RoboDK station: Robot_3_2026.rdk

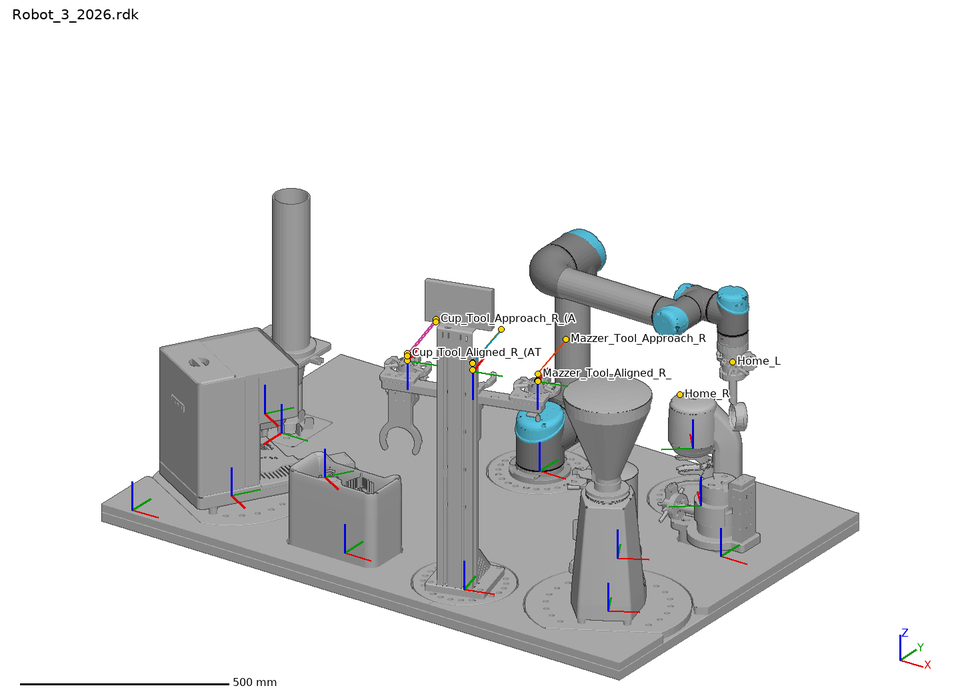
[picture v0: the station drawn from its stored meshes, robots at their saved joint values, targets as dots, program paths as lines]
Station Robot_3_2026 (saved by RoboDK 6.0.6). Poses are relative to the parent item; angles as X-Y-Z fixed-axis rotations.
Station parameters (name, value as stored): IO_5, 1, IO_2, 0, IO_3, 0, IO_4, 0, IO_1, 0, IO_0, 0, 0, 0, 1, 0, 4, 0, 5, 0
  - frame UR5_Base at (0, 0, 0) mm
    - robot UR5: 6 axes
        modified DH rows (alpha deg, a mm, theta deg, d mm): 0, 0, 0, 89.2; 90, 0, 180, 0; 0, 425, 0, 0; 0, 392, 0, 109.3; -90, 0, 0, 94.75; 90, 0, 180, 82.5
        joint limits [-360, -360, -360, -360, -360, -360] to [360, 360, 360, 360, 360, 360]; home [0, -90, -90, 0, 90, 0]; saved at [180, -90, 90, -90, -90, -90]
      - tool Master_Tool_(UR5), TCP at (0, 0, 48.94) mm, size 88.9 x 94.7 x 67.9 mm
      - tool Cup_Tool_Shut_(UR5), TCP at (-34.39, 40.98, 235.56) mm, rotated rx 0 ry 0 rz -50 deg, size 116 x 104.2 x 218.8 mm
      - tool Cup_Tool_Open_(UR5), TCP at (-67.17, 80.05, 235.56) mm, rotated rx 0 ry 0 rz -50 deg, size 166.5 x 104.2 x 218.8 mm
      - tool Mazzer_Tool_(UR5), TCP at (0, 0, 151.76) mm, rotated rx 0 ry 0 rz -50 deg, size 105.5 x 104.2 x 106.6 mm
      - tool Rancilio_Tool_(UR5), TCP at (18.19, -21.68, 194.84) mm, rotated rx 0 ry -3.9 rz -50 deg, size 87.5 x 104.2 x 184.8 mm
      - tool Cup_(UR5), TCP at (-82.31, 98.09, 235.54) mm, rotated rx 0 ry 0 rz -50 deg, size 79 x 78 x 79 mm
    - object UR5_Plate at (0, 0, 0) mm, size 249.9 x 249.9 x 20 mm, geometry from UR5_Plate.STL
    - frame Table_Top at (-700, -700, -20) mm
      - object Table_Top at (0, 0, 0) mm, size 1515 x 1000 x 25 mm, geometry from Table_Top.STL
      - object Table_Cushion at (0, 0, 0) mm, size 1515 x 1000 x 20 mm, geometry from Table_Cushion.STL
      - frame Rancilio at (150, 200, 0) mm, rotated rx 0 ry 0 rz -30 deg
        - object Rancilio at (0, 0, 0) mm, size 399.6 x 458 x 388.3 mm, geometry from Rancilio_Assembly.STL
        - frame Rancilio_Tool at (39.29, 69.7, 222) mm
          - object Rancilio_Tool_Inserted_(Rancilio) at (0, 0, 0) mm, rotated rx 0 ry -90 rz 45 deg, size 87.1 x 104.3 x 184.1 mm, geometry from Rancilio_Tool_Assembly.STL
          - object Rancilio_Tool_Rotated_(Rancilio) at (0, 0, 0) mm, rotated rx 0 ry -90 rz 75 deg, size 87.1 x 104.3 x 184.1 mm, geometry from Rancilio_Tool_Assembly.STL
        - frame Rancilio_Scale at (39, 226.92, 20) mm
          - object Cup_(Rancilio) at (0, -157.52, 65.24) mm, size 79 x 79 x 78 mm, geometry from Supreme_Cup.STL
          - object Rancilio_Scale_Lock at (0, 0, 0) mm, size 100.1 x 260 x 71.4 mm, geometry from Rancilio_Scale_Assembly_1_Lock.STL
          - object Rancilio_Scale_Read at (0, 0, 0) mm, size 100.1 x 260 x 71.4 mm, geometry from Rancilio_Scale_Assembly_1_Read.STL
      - frame Rancilio_Tool_Cleaner at (550, 100, 0) mm
        - object Rancilio_Tool_Cleaner at (0, 0, 0) mm, size 258 x 136.9 x 218.7 mm, geometry from Portafilter_Cleaner_Assembly.STL
      - frame ATI at (900, 100, 0) mm, rotated rx 0 ry 0 rz 15 deg
        - object ATI at (0, 0, 0) mm, size 444.3 x 250 x 843.3 mm, geometry from ATI_Assembly_1.STL
        - frame Cup_Tool_(ATI) at (-164.83, 54.29, 556) mm, rotated rx 180 ry 0 rz 90 deg
          - object Cup_Tool_Shut_(ATI) at (0, 0, 0) mm, size 116 x 104.3 x 218.9 mm, geometry from Cup_Tool_Assembly_Closed.STL
          - target Cup_Tool_Approach_R_(ATI) (Cartesian target) at (200, 0, -20) mm, rotated rx 0 ry 0 rz 50 deg; joints [-77.363, -81.583, -71.578, -116.92, 90.433, -222.544] of UR5
          - target Cup_Tool_Aligned_R_(ATI) (Cartesian target) at (0, 0, -20) mm, rotated rx 0 ry 0 rz 50 deg; joints [-76.522, -110.425, -39.033, -120.623, 90.389, -221.746] of UR5
          - target Cup_Tool_Inserted_R_(ATI) (joint target) at (0, 0, -2) mm, rotated rx 0 ry 0 rz 50 deg; joints [-76.654, -108.705, -44.34, -116.953, 90.001, -221.654] of UR5
          - target Cup_Tool_Mated_R_(ATI) (joint target) at (0, 0, -1) mm, rotated rx 0 ry 0 rz 50 deg; joints [-76.531, -108.58, -44.808, -116.694, 90.407, -221.724] of UR5
          - target Cup_Tool_Attached_R_(ATI) (joint target) at (0, 0, -13) mm, rotated rx 0 ry 0 rz 50 deg; joints [-76.654, -109.734, -41.073, -119.192, 90.001, -221.654] of UR5
          - target Cup_Tool_Rotated_R_(ATI) (joint target) at (0, 0, -13) mm, rotated rx 0 ry 0 rz 140 deg; joints [-76.654, -109.734, -41.073, -119.192, 90.001, -131.654] of UR5
          - target Cup_Tool_Departure_R_(ATI) (joint target) at (200, 0, -13) mm, rotated rx 0 ry 0 rz 140 deg; joints [-77.521, -81.186, -72.909, -115.903, 90.001, -132.521] of UR5
          - target Cup_Tool_Approach_L_(ATI) (joint target) at (200, 0, -20) mm, rotated rx 0 ry 0 rz 50 deg; joints [70.564, -98.372, 71.405, -63.033, -89.998, -254.436] of UR5
          - target Cup_Tool_Aligned_L_(ATI) (joint target) at (0, 0, -20) mm, rotated rx 0 ry 0 rz 50 deg; joints [81.928, -69.509, 38.665, -59.07, -89.569, -243.249] of UR5
          - target Cup_Tool_Inserted_L_(ATI) (joint target) at (0, 0, -2) mm, rotated rx 0 ry 0 rz 50 deg; joints [81.921, -71.276, 44.169, -62.808, -89.552, -243.228] of UR5
          - target Cup_Tool_Mated_L_(ATI) (joint target) at (0, 0, -1) mm, rotated rx 0 ry 0 rz 50 deg; joints [81.836, -71.336, 44.416, -62.995, -89.551, -243.312] of UR5
          - target Cup_Tool_Attached_L_(ATI) (joint target) at (0, 0, -13) mm, rotated rx 0 ry 0 rz 50 deg; joints [81.925, -70.245, 40.897, -60.568, -89.562, -243.241] of UR5
          - target Cup_Tool_Rotated_L_(ATI) (joint target) at (0, 0, -13) mm, rotated rx 0 ry 0 rz 140 deg; joints [81.925, -70.245, 40.897, -60.568, -89.562, -153.241] of UR5
          - target Cup_Tool_Departure_L_(ATI) (joint target) at (200, 0, -13) mm, rotated rx 0 ry 0 rz 140 deg; joints [70.564, -98.814, 72.909, -64.096, -89.998, -164.436] of UR5
        - frame Mazzer_Tool_(ATI) at (165.36, 57.45, 555.5) mm, rotated rx 180 ry 0 rz 90 deg
          - object Mazzer_Tool_(ATI) at (0, 0, 0) mm, size 105.5 x 104.3 x 106.6 mm, geometry from Mazzer_Tool_Assembly.STL
          - target Mazzer_Tool_Approach_R_(ATI) (joint target) at (200, 0, -20) mm, rotated rx 0 ry 0 rz 50 deg; joints [-31.503, -85.319, -68.305, -116.374, 90, -176.503] of UR5
          - target Mazzer_Tool_Aligned_R_(ATI) (joint target) at (0, 0, -20) mm, rotated rx 0 ry 0 rz 50 deg; joints [-45.02, -113.946, -33.907, -122.228, 90.378, -190.259] of UR5
          - target Mazzer_Tool_Inserted_R_(ATI) (joint target) at (-0.58, -1.51, -2.91) mm, rotated rx -0.01 ry -0.4 rz 50.21 deg; joints [-45.095, -111.928, -39.832, -118.239, 90, -190.095] of UR5
          - target Mazzer_Tool_Mated_R_(ATI) (joint target) at (0.03, -0.03, -1.58) mm, rotated rx -0.08 ry -0.01 rz 49.99 deg; joints [-45.032, -111.812, -40.22, -117.969, 90.404, -190.25] of UR5
          - target Mazzer_Tool_Approach_L_(ATI) (joint target) at (200, 0, -20) mm, rotated rx 0 ry 0 rz 50 deg; joints [118.506, -94.678, 68.15, -63.388, -89.525, -206.645] of UR5
          - target Mazzer_Tool_Aligned_L_(ATI) (joint target) at (0, 0, -20) mm, rotated rx 0 ry 0 rz 50 deg; joints [114.077, -65.98, 33.523, -57.458, -89.581, -211.112] of UR5
          - target Mazzer_Tool_Inserted_L_(ATI) (joint target) at (0, 0, -2) mm, rotated rx 0 ry 0 rz 50 deg; joints [114.07, -68.03, 39.626, -61.512, -89.561, -211.089] of UR5
          - target Mazzer_Tool_Mated_L_(ATI) (joint target) at (0, 0, -1) mm, rotated rx 0 ry 0 rz 50 deg; joints [114.069, -68.13, 39.937, -61.723, -89.56, -211.088] of UR5
        - frame Rancilio_Tool_(ATI) at (0.47, 55.43, 555.5) mm, rotated rx 180 ry 0 rz 90 deg
          - object Rancilio_Tool_(ATI) at (0, 0, 0) mm, size 87.5 x 104.3 x 184.8 mm, geometry from Rancilio_Tool_Assembly.STL
          - target Rancilio_Tool_Approach_R_(ATI) (joint target) at (200, 0, -20) mm, rotated rx 0 ry 0 rz 50 deg; joints [-52.246, -78.943, -73.62, -117.435, 90.001, -197.246] of UR5
          - target Rancilio_Tool_Aligned_R_(ATI) (joint target) at (0.2, -0.53, -22.92) mm, rotated rx 0.27 ry -0.38 rz 50.13 deg; joints [-60.08, -108.178, -41.781, -120.208, 89.933, -205.164] of UR5
          - target Rancilio_Tool_Inserted_R_(ATI) (joint target) at (0.24, -0.54, -2.94) mm, rotated rx 0.27 ry -0.38 rz 50.14 deg; joints [-60.089, -106.359, -47.579, -116.227, 89.95, -205.138] of UR5
          - target Rancilio_Tool_Mated_R_(ATI) (joint target) at (0.24, -0.54, -2.94) mm, rotated rx 0.27 ry -0.38 rz 50.14 deg; joints [-60.089, -106.359, -47.579, -116.227, 89.95, -205.138] of UR5
          - target Rancilio_Tool_Approach_L_(ATI) (joint target) at (199.83, 0.84, -20.03) mm, rotated rx -0.01 ry -0.01 rz 49.99 deg; joints [94.213, -101.025, 73.592, -62.577, -89.997, -230.794] of UR5
          - target Rancilio_Tool_Aligned_L_(ATI) (joint target) at (0.22, -0.57, -20.87) mm, rotated rx 0.12 ry -0.38 rz 50.21 deg; joints [97.82, -72.068, 42.273, -60.321, -89.911, -227.136] of UR5
          - target Rancilio_Tool_Inserted_L_(ATI) (joint target) at (0.25, -0.58, -3.24) mm, rotated rx 0.12 ry -0.38 rz 50.21 deg; joints [97.813, -73.65, 47.342, -63.807, -89.894, -227.113] of UR5
          - target Rancilio_Tool_Mated_L_(ATI) (joint target) at (0.25, -0.58, -3.24) mm, rotated rx 0.12 ry -0.38 rz 50.21 deg; joints [97.813, -73.65, 47.342, -63.807, -89.894, -227.113] of UR5
      - frame Mazzer at (1250, 200, 0) mm, rotated rx 0 ry 0 rz 30 deg
        - object Mazzer at (0, 0, 0) mm, size 399.9 x 495 x 614.6 mm, geometry from Mazzer_Assembly_1.STL
        - frame Mazzer_Scale at (0, 250, 20) mm
          - object Rancilio_Tool_(Mazzer) at (0, 40.18, 83.9) mm, rotated rx 0 ry -90 rz 90 deg, size 87.5 x 104.3 x 184.8 mm, geometry from Rancilio_Tool_Assembly.STL
          - object Mazzer_Scale_Lock at (0, 0, 0) mm, size 100.1 x 172.3 x 103.6 mm, geometry from Mazzer_Scale_Assembly_1_Lock.STL
          - object Mazzer_Scale_Read at (0, 0, 0) mm, size 100.1 x 172.3 x 103.6 mm, geometry from Mazzer_Scale_Assembly_1_Read.STL
      - frame Cup_Dispenser at (50, 550, 0) mm, rotated rx 0 ry 0 rz -90 deg
        - object Cup_Dispenser_Shut at (0, 0, 0) mm, size 162 x 208 x 656.6 mm, geometry from Cup_Dispenser_Assembly_Closed.STL
        - object Cup_Dispenser_Open at (0, 0, 0) mm, size 162 x 244.5 x 656.6 mm, geometry from Cup_Dispenser_Assembly_Open.STL
        - object Cup_(Cup_Dispenser) at (0, 27.5, 0) mm, size 79 x 79 x 78 mm, geometry from Supreme_Cup.STL
      - frame PUQ at (1100, 800, 0) mm, rotated rx 0 ry 0 rz 130 deg
        - object PUQ at (0, 0, 0) mm, size 249.7 x 250 x 301 mm, geometry from PUQ_Assembly.STL
        - frame Rancilio_Tool at (0, 18.5, 153.57) mm
          - object Rancilio_Tool_(PUQ) at (0, 0, 0) mm, rotated rx 0 ry -90 rz 90 deg, size 87.1 x 104.3 x 184.1 mm, geometry from Rancilio_Tool_Assembly.STL
      - frame WDT at (1300, 600, 0) mm
        - object Rancilio_Tool_(WDT) at (-10, 0, 133.57) mm, rotated rx 0 ry -90 rz -180 deg, size 87.1 x 104.3 x 184.1 mm, geometry from Rancilio_Tool_Assembly.STL
        - object WDT_Open at (0, 0, 0) mm, size 233 x 150 x 344.6 mm, geometry from UK_Tool_Assembly_Open.STL
        - object WDT_Shut at (0, 0, 0) mm, size 233 x 150 x 244.6 mm, geometry from UK_Tool_Assembly_Shut.STL
      - target Home_R (joint target) at (1186.75, 590.7, 402.76) mm, rotated rx 180 ry 0 rz -40 deg; joints [0, -90, -90, -90, 90, 0] of UR5
      - target Home_L (joint target) at (1186.75, 809.3, 402.76) mm, rotated rx -180 ry 0 rz 0 deg; joints [180, -90, 90, -90, -90, -90] of UR5
  - folder Tool_Programs
    - program Cup_Tool_Attach_R_(ATI) (14 instructions, listed below)
    - program Cup_Tool_Attach_L_(ATI) (14 instructions, listed below)
    - program Cup_Tool_Detach_R_(ATI) (17 instructions, listed below)
    - program Cup_Tool_Detach_L_(ATI) (17 instructions, listed below)
    - program WDT_Open (6 instructions, listed below)
    - program WDT_Shut (6 instructions, listed below)
    - program Mazzer_Tool_Attach_R_(ATI) (12 instructions, listed below)
    - program Mazzer_Tool_Attach_L_(ATI) (12 instructions, listed below)
    - program Mazzer_Tool_Detach_R_(ATI) (16 instructions, listed below)
    - program Mazzer_Tool_Detach_L_(ATI) (16 instructions, listed below)
    - program Rancilio_Tool_Attach_R_(ATI) (12 instructions, listed below)
    - program Rancilio_Tool_Attach_L_(ATI) (12 instructions, listed below)
    - program Rancilio_Tool_Detach_R_(ATI) (15 instructions, listed below)
    - program Rancilio_Tool_Detach_L_(ATI) (15 instructions, listed below)
    - program Cup_Tool_Open_(UR5) (5 instructions, listed below)
    - program Cup_Tool_Shut_(UR5) (5 instructions, listed below)
    - program Student_Tool_Attach (2 instructions, listed below)
    - program Student_Tool_Detach (5 instructions, listed below)
  - folder Visual_Programs
    - program Reset_Simulation_L (25 instructions, listed below)
    - program Reset_Simulation_R (25 instructions, listed below)
    - program Show_Rancilio_Scale_Lock (2 instructions, listed below)
    - program Show_Rancilio_Scale_Read (2 instructions, listed below)
    - program Show_Mazzer_Scale_Lock (2 instructions, listed below)
    - program Show_Mazzer_Scale_Read (2 instructions, listed below)
    - program Show_Mazzer_Scale_Rancilio_Tool (1 instructions, listed below)
    - program Hide_Mazzer_Scale_Rancilio_Tool (1 instructions, listed below)
    - program Show_Rancilio_Scale_Cup (1 instructions, listed below)
    - program Hide_Rancilio_Scale_Cup (1 instructions, listed below)
    - program Show_Cup_Dispenser_Cup (1 instructions, listed below)
    - program Hide_Cup_Dispenser_Cup (1 instructions, listed below)
    - program Show_Cup_Dispenser_Open (2 instructions, listed below)
    - program Show_Cup_Dispenser_Shut (2 instructions, listed below)
    - program Show_WDT_Shut (2 instructions, listed below)
    - program Show_WDT_Open (2 instructions, listed below)
    - program Hide_WDT_Rancilio_Tool (1 instructions, listed below)
    - program Show_WDT_Rancilio_Tool (1 instructions, listed below)
    - program Show_Cup_Tool_Cup (1 instructions, listed below)
    - program Hide_Cup_Tool_Cup (1 instructions, listed below)
    - program Show_Rancilio_Rancilio_Tool_Rotated (1 instructions, listed below)
    - program Hide_Rancilio_Rancilio_Tool_Rotated (1 instructions, listed below)
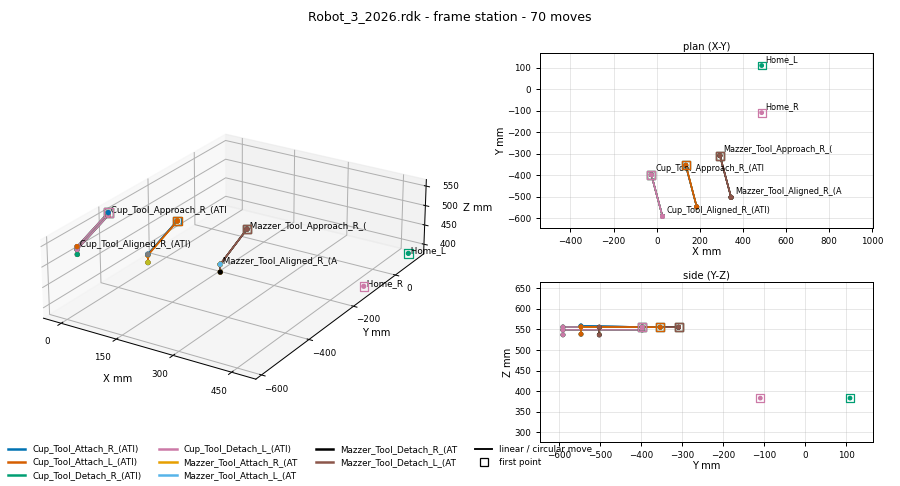
[picture p0: tool path of Robot_3_2026.rdk in frame station, 70 of 70 moves have a stored position in this frame; points joined in program order, loops and branches not executed]

--- program Cup_Tool_Attach_R_(ATI) (robot UR5) ---
  Set Ref.: Cup_Tool_(ATI)
  Set Tool: Master_Tool_(UR5)
  MoveJ (Cup_Tool_Approach_R_(ATI))
  MoveL (Cup_Tool_Aligned_R_(ATI))
  MoveL (Cup_Tool_Mated_R_(ATI))
  Set IO_0=1
  Pause 500 ms
  Hide Cup_Tool_Shut_(ATI)
  Show Cup_Tool_Shut_(UR5)
  MoveL (Cup_Tool_Attached_R_(ATI))
  MoveL (Cup_Tool_Rotated_R_(ATI))
  MoveL (Cup_Tool_Departure_R_(ATI))
  MoveL (Cup_Tool_Approach_R_(ATI))
  Set Ref.: UR5_Base

--- program Cup_Tool_Attach_L_(ATI) (robot UR5) ---
  Set Ref.: Cup_Tool_(ATI)
  Set Tool: Master_Tool_(UR5)
  MoveJ (Cup_Tool_Approach_L_(ATI))
  MoveL (Cup_Tool_Aligned_L_(ATI))
  MoveL (Cup_Tool_Mated_L_(ATI))
  Set IO_0=1
  Pause 500 ms
  Hide Cup_Tool_Shut_(ATI)
  Show Cup_Tool_Shut_(UR5)
  MoveL (Cup_Tool_Attached_L_(ATI))
  MoveL (Cup_Tool_Rotated_L_(ATI))
  MoveL (Cup_Tool_Departure_L_(ATI))
  MoveL (Cup_Tool_Approach_L_(ATI))
  Set Ref.: UR5_Base

--- program Cup_Tool_Detach_R_(ATI) (robot UR5) ---
  Set Ref.: Cup_Tool_(ATI)
  Set Tool: Master_Tool_(UR5)
  MoveJ (Cup_Tool_Approach_R_(ATI))
  MoveL (Cup_Tool_Departure_R_(ATI))
  MoveL (Cup_Tool_Rotated_R_(ATI))
  MoveL (Cup_Tool_Attached_R_(ATI))
  MoveL (Cup_Tool_Mated_R_(ATI))
  Set IO_0=0
  Pause 500 ms
  Set IO_1=1
  Pause 500 ms
  Set IO_1=0
  Hide Cup_Tool_Shut_(UR5)
  Show Cup_Tool_Shut_(ATI)
  MoveL (Cup_Tool_Aligned_R_(ATI))
  MoveL (Cup_Tool_Approach_R_(ATI))
  Set Ref.: UR5_Base

--- program Cup_Tool_Detach_L_(ATI) (robot UR5) ---
  Set Ref.: Cup_Tool_(ATI)
  Set Tool: Master_Tool_(UR5)
  MoveJ (Cup_Tool_Approach_L_(ATI))
  MoveL (Cup_Tool_Departure_L_(ATI))
  MoveL (Cup_Tool_Rotated_L_(ATI))
  MoveL (Cup_Tool_Attached_L_(ATI))
  MoveL (Cup_Tool_Mated_L_(ATI))
  Set IO_0=0
  Pause 500 ms
  Set IO_1=1
  Pause 500 ms
  Set IO_1=0
  Hide Cup_Tool_Shut_(UR5)
  Show Cup_Tool_Shut_(ATI)
  MoveL (Cup_Tool_Aligned_L_(ATI))
  MoveL (Cup_Tool_Approach_L_(ATI))
  Set Ref.: UR5_Base

--- program WDT_Open (robot UR5) ---
  Set IO_4=1
  Pause 500 ms
  Set IO_4=0
  Pause 500 ms
  Hide WDT_Shut
  Show WDT_Open

--- program WDT_Shut (robot UR5) ---
  Set IO_5=1
  Pause 500 ms
  Set IO_5=0
  Pause 500 ms
  Hide WDT_Open
  Show WDT_Shut

--- program Mazzer_Tool_Attach_R_(ATI) (robot UR5) ---
  Set Ref.: Mazzer_Tool_(ATI)
  Set Tool: Master_Tool_(UR5)
  MoveJ (Mazzer_Tool_Approach_R_(ATI))
  MoveL (Mazzer_Tool_Aligned_R_(ATI))
  MoveL (Mazzer_Tool_Mated_R_(ATI))
  Set IO_0=1
  Pause 500 ms
  Hide Mazzer_Tool_(ATI)
  Show Mazzer_Tool_(UR5)
  MoveL (Mazzer_Tool_Aligned_R_(ATI))
  MoveL (Mazzer_Tool_Approach_R_(ATI))
  Set Ref.: UR5_Base

--- program Mazzer_Tool_Attach_L_(ATI) (robot UR5) ---
  Set Ref.: Mazzer_Tool_(ATI)
  Set Tool: Master_Tool_(UR5)
  MoveJ (Mazzer_Tool_Approach_L_(ATI))
  MoveL (Mazzer_Tool_Aligned_L_(ATI))
  MoveL (Mazzer_Tool_Mated_L_(ATI))
  Set IO_0=1
  Pause 500 ms
  Hide Mazzer_Tool_(ATI)
  Show Mazzer_Tool_(UR5)
  MoveL (Mazzer_Tool_Aligned_L_(ATI))
  MoveL (Mazzer_Tool_Approach_L_(ATI))
  Set Ref.: UR5_Base

--- program Mazzer_Tool_Detach_R_(ATI) (robot UR5) ---
  Set Ref.: Mazzer_Tool_(ATI)
  Set Tool: Master_Tool_(UR5)
  MoveJ (Mazzer_Tool_Approach_R_(ATI))
  MoveL (Mazzer_Tool_Aligned_R_(ATI))
  MoveL (Mazzer_Tool_Mated_R_(ATI))
  Set IO_0=0
  Pause 500 ms
  Set IO_1=1
  Pause 500 ms
  Set IO_1=0
  Hide Mazzer_Tool_(UR5)
  Show Mazzer_Tool_(ATI)
  MoveL (Mazzer_Tool_Aligned_R_(ATI))
  MoveL (Mazzer_Tool_Approach_R_(ATI))
  Set Ref.: UR5_Base
  Set Tool: Master_Tool_(UR5)

--- program Mazzer_Tool_Detach_L_(ATI) (robot UR5) ---
  Set Ref.: Mazzer_Tool_(ATI)
  Set Tool: Master_Tool_(UR5)
  MoveJ (Mazzer_Tool_Approach_L_(ATI))
  MoveL (Mazzer_Tool_Aligned_L_(ATI))
  MoveL (Mazzer_Tool_Mated_L_(ATI))
  Set IO_0=0
  Pause 500 ms
  Set IO_1=1
  Pause 500 ms
  Set IO_1=0
  Hide Mazzer_Tool_(UR5)
  Show Mazzer_Tool_(ATI)
  MoveL (Mazzer_Tool_Aligned_L_(ATI))
  MoveL (Mazzer_Tool_Approach_L_(ATI))
  Set Ref.: UR5_Base
  Set Tool: Master_Tool_(UR5)

--- program Rancilio_Tool_Attach_R_(ATI) (robot UR5) ---
  Set Ref.: Rancilio_Tool_(ATI)
  Set Tool: Master_Tool_(UR5)
  MoveJ (Rancilio_Tool_Approach_R_(ATI))
  MoveL (Rancilio_Tool_Aligned_R_(ATI))
  MoveL (Rancilio_Tool_Mated_R_(ATI))
  Set IO_0=1
  Pause 500 ms
  Hide Rancilio_Tool_(ATI)
  Show Rancilio_Tool_(UR5)
  MoveL (Rancilio_Tool_Aligned_R_(ATI))
  MoveL (Rancilio_Tool_Approach_R_(ATI))
  Set Ref.: UR5_Base

--- program Rancilio_Tool_Attach_L_(ATI) (robot UR5) ---
  Set Ref.: Rancilio_Tool_(ATI)
  Set Tool: Master_Tool_(UR5)
  MoveJ (Rancilio_Tool_Approach_L_(ATI))
  MoveL (Rancilio_Tool_Aligned_L_(ATI))
  MoveL (Rancilio_Tool_Mated_L_(ATI))
  Set IO_0=1
  Pause 500 ms
  Hide Rancilio_Tool_(ATI)
  Show Rancilio_Tool_(UR5)
  MoveL (Rancilio_Tool_Aligned_L_(ATI))
  MoveL (Rancilio_Tool_Approach_L_(ATI))
  Set Ref.: UR5_Base

--- program Rancilio_Tool_Detach_R_(ATI) (robot UR5) ---
  Set Ref.: Rancilio_Tool_(ATI)
  Set Tool: Master_Tool_(UR5)
  MoveJ (Rancilio_Tool_Approach_R_(ATI))
  MoveL (Rancilio_Tool_Aligned_R_(ATI))
  MoveL (Rancilio_Tool_Mated_R_(ATI))
  Set IO_0=0
  Pause 500 ms
  Set IO_1=1
  Pause 500 ms
  Set IO_1=0
  Hide Rancilio_Tool_(UR5)
  Show Rancilio_Tool_(ATI)
  MoveL (Rancilio_Tool_Aligned_R_(ATI))
  MoveL (Rancilio_Tool_Approach_R_(ATI))
  Set Ref.: UR5_Base

--- program Rancilio_Tool_Detach_L_(ATI) (robot UR5) ---
  Set Ref.: Rancilio_Tool_(ATI)
  Set Tool: Master_Tool_(UR5)
  MoveJ (Rancilio_Tool_Approach_L_(ATI))
  MoveL (Rancilio_Tool_Aligned_L_(ATI))
  MoveL (Rancilio_Tool_Mated_L_(ATI))
  Set IO_0=0
  Pause 500 ms
  Set IO_1=1
  Pause 500 ms
  Set IO_1=0
  Hide Rancilio_Tool_(UR5)
  Show Rancilio_Tool_(ATI)
  MoveL (Rancilio_Tool_Aligned_L_(ATI))
  MoveL (Rancilio_Tool_Approach_L_(ATI))
  Set Ref.: UR5_Base

--- program Cup_Tool_Open_(UR5) (robot UR5) ---
  Set IO_2=1
  Hide Cup_Tool_Shut_(UR5)
  Show Cup_Tool_Open_(UR5)
  Pause 500 ms
  Set IO_2=0

--- program Cup_Tool_Shut_(UR5) (robot UR5) ---
  Set IO_3=1
  Hide Cup_Tool_Open_(UR5)
  Show Cup_Tool_Shut_(UR5)
  Pause 500 ms
  Set IO_3=0

--- program Student_Tool_Attach (robot UR5) ---
  Set IO_0=1
  Pause 500 ms

--- program Student_Tool_Detach (robot UR5) ---
  Set IO_0=0
  Pause 500 ms
  Set IO_1=1
  Pause 500 ms
  Set IO_1=0

--- program Reset_Simulation_L (robot UR5) ---
  MoveJ (Home_L)
  Show Master_Tool_(UR5)
  Hide Cup_Tool_Shut_(UR5)
  Hide Cup_Tool_Open_(UR5)
  Hide Mazzer_Tool_(UR5)
  Hide Rancilio_Tool_(UR5)
  Hide Cup_(UR5)
  Hide Rancilio_Tool_Inserted_(Rancilio)
  Hide Rancilio_Tool_Rotated_(Rancilio)
  Hide Cup_(Rancilio)
  Hide Rancilio_Scale_Read
  Show Rancilio_Scale_Lock
  Show Cup_Tool_Shut_(ATI)
  Show Mazzer_Tool_(ATI)
  Show Rancilio_Tool_(ATI)
  Hide Mazzer_Scale_Read
  Show Mazzer_Scale_Lock
  Hide Cup_Dispenser_Open
  Show Cup_Dispenser_Shut
  Hide Cup_(Cup_Dispenser)
  Hide Rancilio_Tool_(PUQ)
  Hide Rancilio_Tool_(Mazzer)
  Hide WDT_Open
  Show WDT_Shut
  Hide Rancilio_Tool_(WDT)

--- program Reset_Simulation_R (robot UR5) ---
  MoveJ (Home_R)
  Show Master_Tool_(UR5)
  Hide Cup_Tool_Shut_(UR5)
  Hide Cup_Tool_Open_(UR5)
  Hide Mazzer_Tool_(UR5)
  Hide Rancilio_Tool_(UR5)
  Hide Cup_(UR5)
  Hide Rancilio_Tool_Inserted_(Rancilio)
  Hide Rancilio_Tool_Rotated_(Rancilio)
  Hide Cup_(Rancilio)
  Hide Rancilio_Scale_Read
  Show Rancilio_Scale_Lock
  Show Cup_Tool_Shut_(ATI)
  Show Mazzer_Tool_(ATI)
  Show Rancilio_Tool_(ATI)
  Hide Mazzer_Scale_Read
  Show Mazzer_Scale_Lock
  Hide Cup_Dispenser_Open
  Show Cup_Dispenser_Shut
  Hide Cup_(Cup_Dispenser)
  Hide Rancilio_Tool_(PUQ)
  Hide Rancilio_Tool_(Mazzer)
  Hide WDT_Open
  Show WDT_Shut
  Hide Rancilio_Tool_(WDT)

--- program Show_Rancilio_Scale_Lock (robot UR5) ---
  Show Rancilio_Scale_Lock
  Hide Rancilio_Scale_Read

--- program Show_Rancilio_Scale_Read (robot UR5) ---
  Hide Rancilio_Scale_Lock
  Show Rancilio_Scale_Read

--- program Show_Mazzer_Scale_Lock (robot UR5) ---
  Hide Mazzer_Scale_Read
  Show Mazzer_Scale_Lock

--- program Show_Mazzer_Scale_Read (robot UR5) ---
  Hide Mazzer_Scale_Lock
  Show Mazzer_Scale_Read

--- program Show_Mazzer_Scale_Rancilio_Tool (robot UR5) ---
  Show Rancilio_Tool_(Mazzer)

--- program Hide_Mazzer_Scale_Rancilio_Tool (robot UR5) ---
  Hide Rancilio_Tool_(Mazzer)

--- program Show_Rancilio_Scale_Cup (robot UR5) ---
  Show Cup_(Rancilio)

--- program Hide_Rancilio_Scale_Cup (robot UR5) ---
  Hide Cup_(Rancilio)

--- program Show_Cup_Dispenser_Cup (robot UR5) ---
  Show Cup_(Cup_Dispenser)

--- program Hide_Cup_Dispenser_Cup (robot UR5) ---
  Hide Cup_(Cup_Dispenser)

--- program Show_Cup_Dispenser_Open (robot UR5) ---
  Hide Cup_Dispenser_Shut
  Show Cup_Dispenser_Open

--- program Show_Cup_Dispenser_Shut (robot UR5) ---
  Hide Cup_Dispenser_Open
  Show Cup_Dispenser_Shut

--- program Show_WDT_Shut (robot UR5) ---
  Hide WDT_Open
  Show WDT_Shut

--- program Show_WDT_Open (robot UR5) ---
  Hide WDT_Shut
  Show WDT_Open

--- program Hide_WDT_Rancilio_Tool (robot UR5) ---
  Hide Rancilio_Tool_(WDT)

--- program Show_WDT_Rancilio_Tool (robot UR5) ---
  Show Rancilio_Tool_(WDT)

--- program Show_Cup_Tool_Cup (robot UR5) ---
  Show Cup_(UR5)

--- program Hide_Cup_Tool_Cup (robot UR5) ---
  Hide Cup_(UR5)

--- program Show_Rancilio_Rancilio_Tool_Rotated (robot UR5) ---
  Show Rancilio_Tool_Rotated_(Rancilio)

--- program Hide_Rancilio_Rancilio_Tool_Rotated (robot UR5) ---
  Hide Rancilio_Tool_Rotated_(Rancilio)
